RoboDK station: RoboDK Simulation.rdk

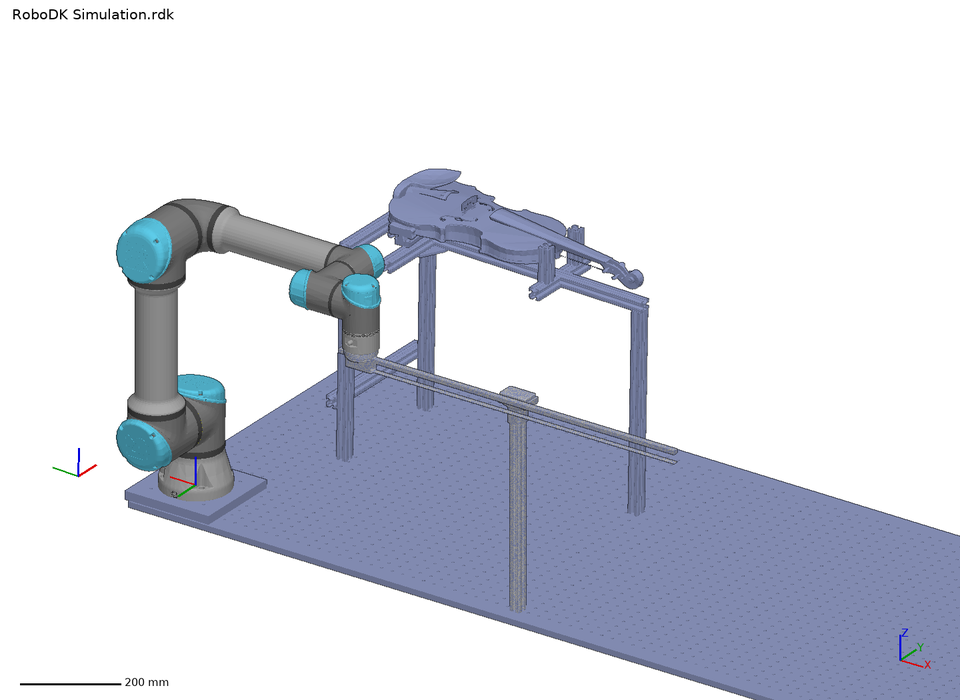
[picture v0: the station drawn from its stored meshes, robots at their saved joint values, targets as dots, program paths as lines]
Station RoboDK Simulation (saved by RoboDK 6.0.4). Poses are relative to the parent item; angles as X-Y-Z fixed-axis rotations.
  - frame UR7e Base at (0, 1428.5, 0) mm, rotated rx 0 ry 0 rz -179.82 deg
    - robot UR7e: 6 axes, payload 5 kg, reach 850 mm, repeatability 0.03 mm, weight 18.4 kg
        modified DH rows (alpha deg, a mm, theta deg, d mm): 0, 0, 0, 162.5; 90, 0, 180, 0; 0, 425, 0, 0; 0, 392.25, 0, 133.3; -90, 0, 0, 99.7; 90, 0, 180, 99.6
        joint limits [-360, -360, -360, -360, -360, -360] to [360, 360, 360, 360, 360, 360]; home [0, -90, -90, 0, 90, 0]; saved at [180, -90, -90, -90, 90, 90]
      - tool UR7e_ToolFlange, TCP at (0, 0, 200) mm, size 812.5 x 69.3 x 45.1 mm, geometry from UR7e_ToolFlange.step
    - object UR7e_Base at (0, 0, 0) mm, size 203.2 x 203.2 x 19 mm, geometry from UR7e_Base.step
  - frame Frame 2 at (415.7, 428.5, 535) mm, rotated rx 1.08 ry 0 rz 90 deg
    - object ViolinFixture at (0, 0, 0) mm, size 330.2 x 660.4 x 582.9 mm, geometry from ViolinFixture.step
  - frame Frame 3 at (-64, -64, -20) mm
    - object OpticalTable at (0, -1958, -32) mm, size 1949.2 x 819.7 x 12.7 mm, geometry from OpticalTable.step
    - object RosinHolder at (0, 0, 0) mm, size 69.8 x 44.4 x 480.5 mm, geometry from RosinHolder.step
